// TIA Portal V21 export
DATA_BLOCK "HMI_Zustand_DB"   // DB6
{ S7_Optimized_Access := 'TRUE' }
// stored: MemoryReserve 100
   VAR
      state : Int;
      einschubachse_einfahren_enabled : Bool;   // Bedingungen für einfahren der Einschubachse sind erfüllt
      Ref_enabled : Bool;   // Bedingungen für Referenzierung sind erfüllt
      jog_mode_enabled : Bool;   // Bedingungen für jog-mode erfüllt
      absolut_pos_enabled : Bool;   // Bedingungen für absolut-pos erfüllt
      relativ_pos_enabled : Bool;   // Bedingungen für relativ-pos erfüllt
      magazinieren_enabled : Bool;   // Bedingungen für magazinieren erfüllt
      abholen_enabeld : Bool;   // Bedingungen für abholen erfüllt
      ref_mode : Bool;   // Referenzierung aktiv
      einschubachse_mode : Bool;   // Einschubachse einfahren aktiv
      jog_mode : Bool;   // jog-mode aktiv
      absolut_pos : Bool;   // absolut-pos aktiv
      relativ_pos : Bool;   // relativ-pos aktiv
      magazinieren : Bool;   // magazinieren aktiv
      abholen : Bool;   // abholen aktiv
      AxisRef_all : Bool;   // Alle Achsen sind referenziert
      Einschubachse_eingefahren : Bool;   // Einschubachse ist eingefahren
      ActPos_absoult_h : LReal;   // angepasste Position für horizontae Achse in [cm]
      ActPos_absoult_v : LReal;   // angepasste Position für vertikale Achse in [cm]
      ActPos_animation_h : Int;   // Wert für Animatio der horizobtalen Achsen
      ActPos_animation_v : Int;   // Wert für Animation der vertikalen Achsen
      AxisEnabled_h : Bool;
      AxisPosOK_h : Bool;
      AxisRef_h : Bool;
      AxisError_h : Bool;
      Error_h : Bool;
      ActVel_h : LReal;
      ActPos_h : LReal;
      AxisEnabled_v : Bool;
      AxisPosOK_v : Bool;
      AxisRef_v : Bool;
      AxisError_v : Bool;
      Error_v : Bool;
      ActVel_v : LReal;
      ActPos_v : LReal;
      AxisRef_z : Bool;
      Error_z : Bool;
      AxisEnabled_z : Bool;
      ErrorID_z : Word;
      ActVel_z : LReal;
      ActPos_z : LReal;
   END_VAR
BEGIN
END_DATA_BLOCK
